(* IEC 61131-3 sources: plc-ci-toolkit/ci/tests/samples/sa_probe_src/src/POUs/FB_SaSkip, 1 file *)

(* ---- FB_SaSkip.decl.st ---- *)
// Назначение: зонд статанализа — объект без анализа
{attribute 'no-analysis'}
FUNCTION_BLOCK FB_SaSkip
VAR_INPUT
    xIn : BOOL;
END_VAR
VAR
    iSkippedUnused : INT;           // SA0033 не должно быть: no-analysis
END_VAR
